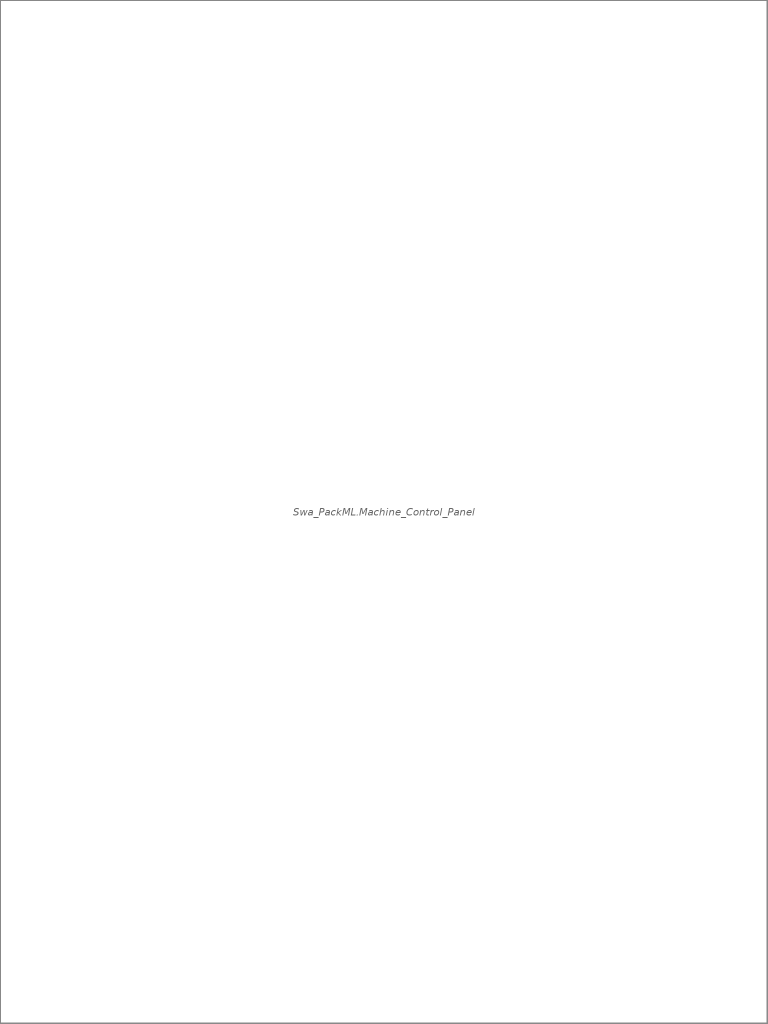
VISUALIZATION Visualization  // 768x1024
    Frame (0,0 768x1024)
        shows Swa_PackML.Machine_Control_Panel(AlarmAdmin := MAIN.Machine.alarmAdmin, ModuleSelector := MAIN.Machine.moduleSelector)
END_VISUALIZATION

(* stored: Version 1.1.0.1, ProductVersion 3.1.4024.12
   Visu Visualization: Id {5b1a45dc-707a-4846-a3d6-72a242e82b9a} *)
